FUNCTION_BLOCK PutWorkpiece (* Basic Function Block Type *)
  (* Standard: 61499-2 *)
  (* Version 0.0, 7/2/2026, Template *)
  PACKAGE Main;
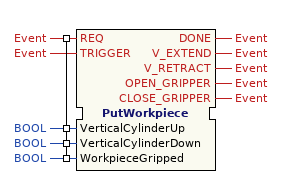
  EVENT_INPUT
    REQ WITH VerticalCylinderUp, VerticalCylinderDown, WorkpieceGripped; (* Normal Execution Request *)
    TRIGGER;
  END_EVENT
  EVENT_OUTPUT
    DONE; (* Initialization Confirm *)
    V_EXTEND; (* Execution Confirmation *)
    V_RETRACT;
    OPEN_GRIPPER;
    CLOSE_GRIPPER;
  END_EVENT
  VAR_INPUT
    VerticalCylinderUp : BOOL; (* Input event qualifier *)
    VerticalCylinderDown : BOOL;
    WorkpieceGripped : BOOL;
  END_VAR
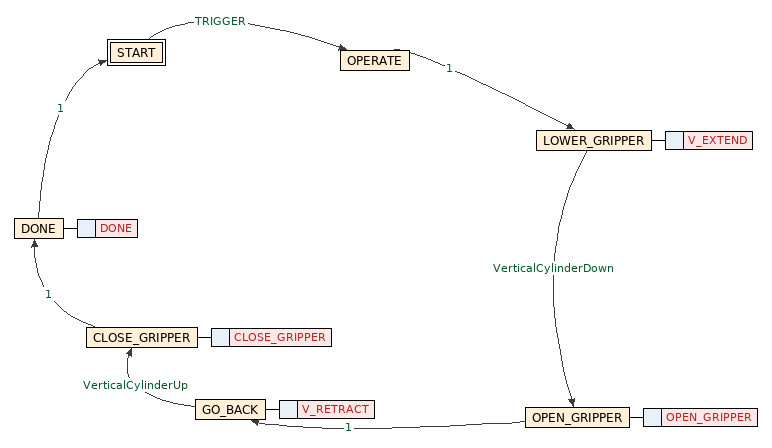
  EC_STATES
    START; (* Initial State *)
    OPERATE;
    LOWER_GRIPPER : -> V_EXTEND;
    OPEN_GRIPPER : -> OPEN_GRIPPER;
    GO_BACK : -> V_RETRACT;
    CLOSE_GRIPPER : -> CLOSE_GRIPPER;
    DONE : -> DONE;
  END_STATES
  EC_TRANSITIONS
    START TO OPERATE := TRIGGER;
    OPERATE TO LOWER_GRIPPER := 1;
    LOWER_GRIPPER TO OPEN_GRIPPER := VerticalCylinderDown;
    OPEN_GRIPPER TO GO_BACK := 1;
    GO_BACK TO CLOSE_GRIPPER := VerticalCylinderUp;
    CLOSE_GRIPPER TO DONE := 1;
    DONE TO START := 1;
  END_TRANSITIONS
  ALGORITHM INIT IN ST: (* Initialization algorithm *)
;
  END_ALGORITHM
  ALGORITHM REQ IN ST: (* Normally executed algorithm *)
;
  END_ALGORITHM
END_FUNCTION_BLOCK
